FUNCTION_BLOCK EPUCK_PROX (* E-puck sensors reading *)
  (* Standard: 61499-2; Classification: SIFB; ApplicationDomain: Robotics; Function: Sensor; Type: SIFB; Description: PROX0..PROX7 gross values *)
  (* Version 1.0, 2026-10-22, Mauricio Martins Taques Filho, GASR/UDESC, Initial version *)
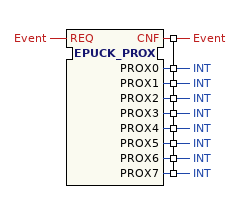
  EVENT_INPUT
    REQ; (* Request a input *)
  END_EVENT
  EVENT_OUTPUT
    CNF WITH PROX0, PROX1, PROX2, PROX3, PROX4, PROX5, PROX6, PROX7; (* Input ready *)
  END_EVENT
  VAR_OUTPUT
    PROX0 : INT; (* Upper right sensor *)
    PROX1 : INT; (* Right/Front sensor *)
    PROX2 : INT; (* Right sensor *)
    PROX3 : INT; (* Right/Back sensor *)
    PROX4 : INT; (* Left/Back sensor *)
    PROX5 : INT; (* Left sensor *)
    PROX6 : INT; (* Left/Front sensor *)
    PROX7 : INT; (* Upper left sensor *)
  END_VAR
  SERVICE APPLICATION/RESOURCE
    SEQUENCE Read
      APPLICATION.REQ() -> APPLICATION.CNF(PROX0,PROX1,PROX2,PROX3,PROX4,PROX5,PROX6,PROX7);
    END_SEQUENCE
  END_SERVICE
END_FUNCTION_BLOCK
